Staubli VAL3: bind.pgx

program bind()
  local string l_slbl
  local num l_i
begin
  userPageBindClick("safepoint","btnback",bBack,true)
  userPageBindClick("safepoint","btn1",bTeach,true)
  userPageBindClick("safepoint","btn2",bMove,true)

  userPageBind("safepoint","lst1","options",sList,size(sList),"r")
  userPageBind("safepoint","lst1","value",sSelPoint,1,"rw")

  userPageBind("safepoint","chk1","checked",bActive,1,"rw")

  for l_i = 0 to 5
    l_slbl="lbl3"+toString("",l_i)
    userPageBind("safepoint",l_slbl,"innerHTML",sTRSF[l_i],1,"r")
  endFor
end
